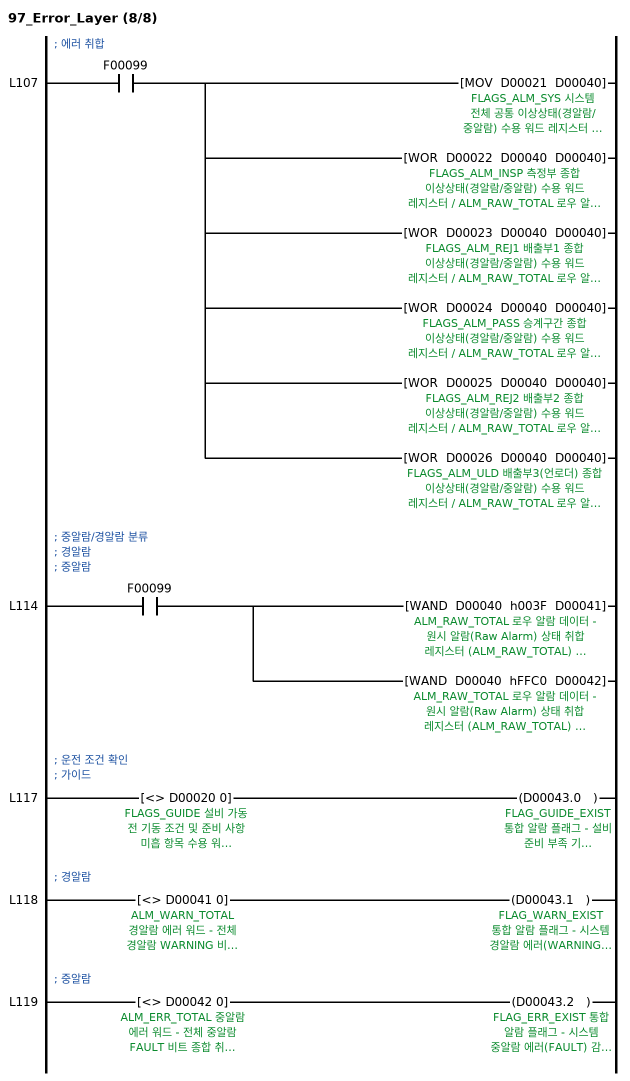
[picture p24: 97_Error_Layer rungs L107-L119]
// 에러 취합
; L107
LOAD      F00099
MOV       D00021 D00040	// FLAGS_ALM_SYS 시스템 전체 공통 이상상태(경알람/중알람) 수용 워드 레지스터 / ALM_RAW_TOTAL 로우 알람 데이터 - 원시 알람(Raw Alarm) 상태 취합 레지스터 (ALM_RAW_TOTAL)
WOR       D00022 D00040 D00040	// FLAGS_ALM_INSP 측정부 종합 이상상태(경알람/중알람) 수용 워드 레지스터 / ALM_RAW_TOTAL 로우 알람 데이터 - 원시 알람(Raw Alarm) 상태 취합 레지스터 (ALM_RAW_TOTAL) / ALM_RAW_TOTAL 로우 알람 데이터 - 원시 알람(Raw Alarm) 상태 취합 레지스터 (ALM_RAW_TOTAL)
WOR       D00023 D00040 D00040	// FLAGS_ALM_REJ1 배출부1 종합 이상상태(경알람/중알람) 수용 워드 레지스터 / ALM_RAW_TOTAL 로우 알람 데이터 - 원시 알람(Raw Alarm) 상태 취합 레지스터 (ALM_RAW_TOTAL) / ALM_RAW_TOTAL 로우 알람 데이터 - 원시 알람(Raw Alarm) 상태 취합 레지스터 (ALM_RAW_TOTAL)
WOR       D00024 D00040 D00040	// FLAGS_ALM_PASS 승계구간 종합 이상상태(경알람/중알람) 수용 워드 레지스터 / ALM_RAW_TOTAL 로우 알람 데이터 - 원시 알람(Raw Alarm) 상태 취합 레지스터 (ALM_RAW_TOTAL) / ALM_RAW_TOTAL 로우 알람 데이터 - 원시 알람(Raw Alarm) 상태 취합 레지스터 (ALM_RAW_TOTAL)
WOR       D00025 D00040 D00040	// FLAGS_ALM_REJ2 배출부2 종합 이상상태(경알람/중알람) 수용 워드 레지스터 / ALM_RAW_TOTAL 로우 알람 데이터 - 원시 알람(Raw Alarm) 상태 취합 레지스터 (ALM_RAW_TOTAL) / ALM_RAW_TOTAL 로우 알람 데이터 - 원시 알람(Raw Alarm) 상태 취합 레지스터 (ALM_RAW_TOTAL)
WOR       D00026 D00040 D00040	// FLAGS_ALM_ULD 배출부3(언로더) 종합 이상상태(경알람/중알람) 수용 워드 레지스터 / ALM_RAW_TOTAL 로우 알람 데이터 - 원시 알람(Raw Alarm) 상태 취합 레지스터 (ALM_RAW_TOTAL) / ALM_RAW_TOTAL 로우 알람 데이터 - 원시 알람(Raw Alarm) 상태 취합 레지스터 (ALM_RAW_TOTAL)
// 중알람/경알람 분류
; L114
LOAD      F00099
WAND      D00040 h003F D00041	// ALM_RAW_TOTAL 로우 알람 데이터 - 원시 알람(Raw Alarm) 상태 취합 레지스터 (ALM_RAW_TOTAL) / ALM_WARN_TOTAL 경알람 에러 워드 - 전체 경알람 WARNING 비트 종합 취합 레지스터 (ALM_WARN_TOTAL)
WAND      D00040 hFFC0 D00042	// ALM_RAW_TOTAL 로우 알람 데이터 - 원시 알람(Raw Alarm) 상태 취합 레지스터 (ALM_RAW_TOTAL) / ALM_ERR_TOTAL 중알람 에러 워드 - 전체 중알람 FAULT 비트 종합 취합 레지스터 (ALM_ERR_TOTAL)
// output comment: 경알람
// output comment: 중알람
// 운전 조건 확인
; L117
LOAD<>    D00020 0	// FLAGS_GUIDE 설비 가동 전 기동 조건 및 준비 사항 미흡 항목 수용 워드 레지스터
OUT       D00043.0	// FLAG_GUIDE_EXIST 통합 알람 플래그 - 설비 준비 부족 기동 불허(GUIDE) 활성화
// output comment: 가이드
; L118
LOAD<>    D00041 0	// ALM_WARN_TOTAL 경알람 에러 워드 - 전체 경알람 WARNING 비트 종합 취합 레지스터 (ALM_WARN_TOTAL)
OUT       D00043.1	// FLAG_WARN_EXIST 통합 알람 플래그 - 시스템 경알람 에러(WARNING) 감지 활성화
// output comment: 경알람
; L119
LOAD<>    D00042 0	// ALM_ERR_TOTAL 중알람 에러 워드 - 전체 중알람 FAULT 비트 종합 취합 레지스터 (ALM_ERR_TOTAL)
OUT       D00043.2	// FLAG_ERR_EXIST 통합 알람 플래그 - 시스템 중알람 에러(FAULT) 감지 활성화
// output comment: 중알람

PROGRAM 98_Output_Layer (task: 스캔 프로그램)

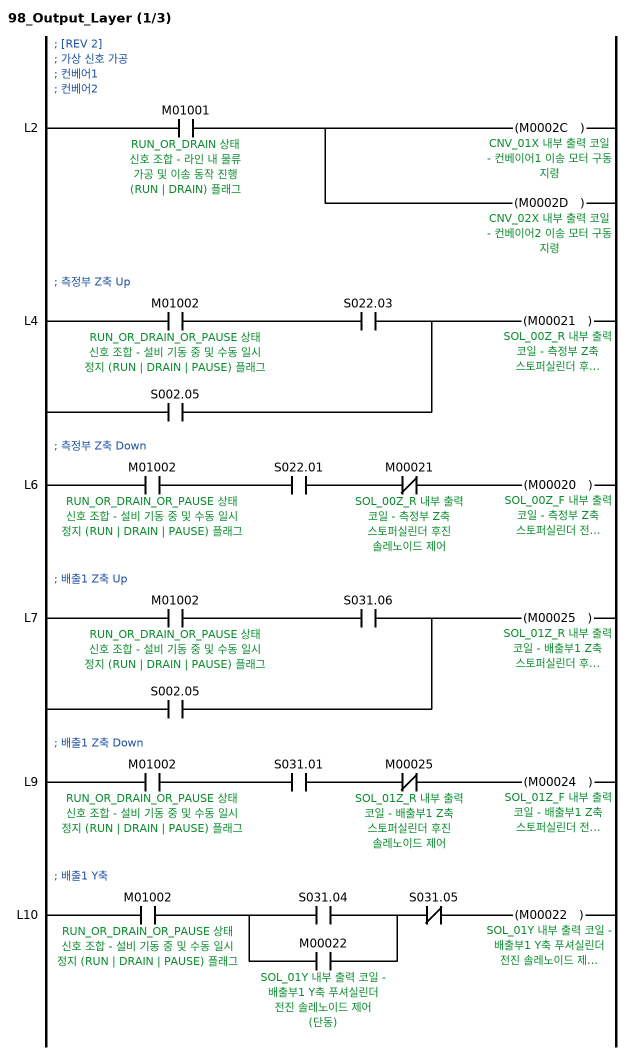
// [REV 2]
// 가상 신호 가공
; L2
LOAD      M01001	// RUN_OR_DRAIN 상태 신호 조합 - 라인 내 물류 가공 및 이송 동작 진행 (RUN | DRAIN) 플래그
OUT       M0002C	// CNV_01X 내부 출력 코일 - 컨베이어1 이송 모터 구동 지령
OUT       M0002D	// CNV_02X 내부 출력 코일 - 컨베이어2 이송 모터 구동 지령
// output comment: 컨베어1
// output comment: 컨베어2
; L4
LOAD      M01002	// RUN_OR_DRAIN_OR_PAUSE 상태 신호 조합 - 설비 기동 중 및 수동 일시 정지 (RUN | DRAIN | PAUSE) 플래그
AND       S022.03
OR        S002.05
OUT       M00021	// SOL_00Z_R 내부 출력 코일 - 측정부 Z축 스토퍼실린더 후진 솔레노이드 제어
// output comment: 측정부 Z축 Up
; L6
LOAD      M01002	// RUN_OR_DRAIN_OR_PAUSE 상태 신호 조합 - 설비 기동 중 및 수동 일시 정지 (RUN | DRAIN | PAUSE) 플래그
AND       S022.01
AND NOT   M00021	// SOL_00Z_R 내부 출력 코일 - 측정부 Z축 스토퍼실린더 후진 솔레노이드 제어
OUT       M00020	// SOL_00Z_F 내부 출력 코일 - 측정부 Z축 스토퍼실린더 전진 솔레노이드 제어
// output comment: 측정부 Z축 Down
; L7
LOAD      M01002	// RUN_OR_DRAIN_OR_PAUSE 상태 신호 조합 - 설비 기동 중 및 수동 일시 정지 (RUN | DRAIN | PAUSE) 플래그
AND       S031.06
OR        S002.05
OUT       M00025	// SOL_01Z_R 내부 출력 코일 - 배출부1 Z축 스토퍼실린더 후진 솔레노이드 제어
// output comment: 배출1 Z축 Up
; L9
LOAD      M01002	// RUN_OR_DRAIN_OR_PAUSE 상태 신호 조합 - 설비 기동 중 및 수동 일시 정지 (RUN | DRAIN | PAUSE) 플래그
AND       S031.01
AND NOT   M00025	// SOL_01Z_R 내부 출력 코일 - 배출부1 Z축 스토퍼실린더 후진 솔레노이드 제어
OUT       M00024	// SOL_01Z_F 내부 출력 코일 - 배출부1 Z축 스토퍼실린더 전진 솔레노이드 제어
// output comment: 배출1 Z축 Down
; L10
LOAD      M01002	// RUN_OR_DRAIN_OR_PAUSE 상태 신호 조합 - 설비 기동 중 및 수동 일시 정지 (RUN | DRAIN | PAUSE) 플래그
LOAD      S031.04
OR        M00022	// SOL_01Y 내부 출력 코일 - 배출부1 Y축 푸셔실린더 전진 솔레노이드 제어 (단동)
AND LOAD
AND NOT   S031.05
OUT       M00022	// SOL_01Y 내부 출력 코일 - 배출부1 Y축 푸셔실린더 전진 솔레노이드 제어 (단동)
// output comment: 배출1 Y축

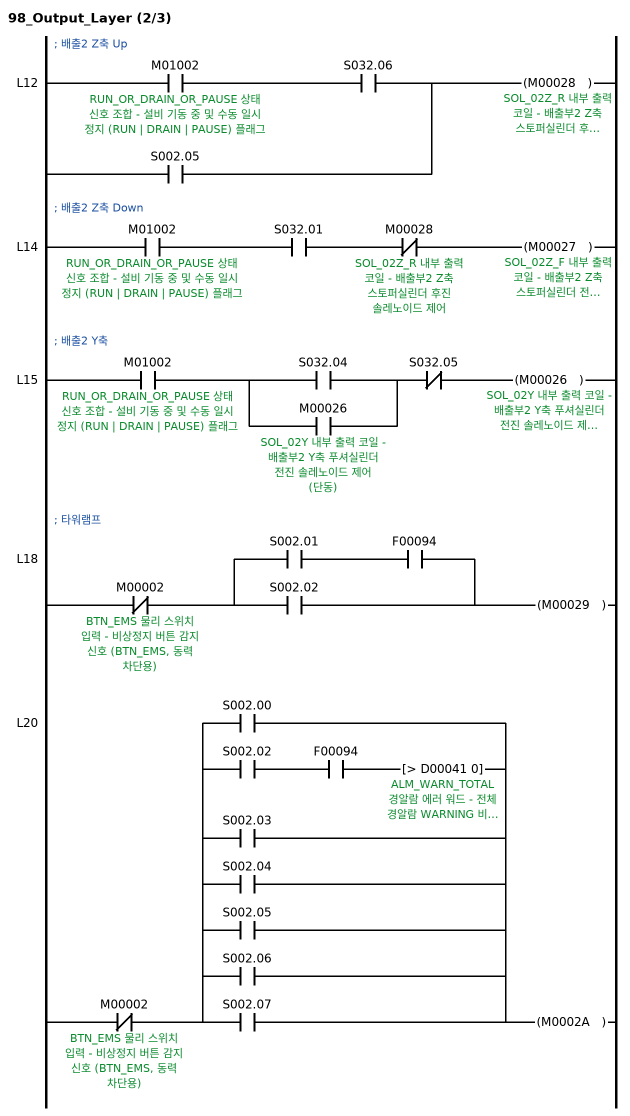
; L12
LOAD      M01002	// RUN_OR_DRAIN_OR_PAUSE 상태 신호 조합 - 설비 기동 중 및 수동 일시 정지 (RUN | DRAIN | PAUSE) 플래그
AND       S032.06
OR        S002.05
OUT       M00028	// SOL_02Z_R 내부 출력 코일 - 배출부2 Z축 스토퍼실린더 후진 솔레노이드 제어
// output comment: 배출2 Z축 Up
; L14
LOAD      M01002	// RUN_OR_DRAIN_OR_PAUSE 상태 신호 조합 - 설비 기동 중 및 수동 일시 정지 (RUN | DRAIN | PAUSE) 플래그
AND       S032.01
AND NOT   M00028	// SOL_02Z_R 내부 출력 코일 - 배출부2 Z축 스토퍼실린더 후진 솔레노이드 제어
OUT       M00027	// SOL_02Z_F 내부 출력 코일 - 배출부2 Z축 스토퍼실린더 전진 솔레노이드 제어
// output comment: 배출2 Z축 Down
; L15
LOAD      M01002	// RUN_OR_DRAIN_OR_PAUSE 상태 신호 조합 - 설비 기동 중 및 수동 일시 정지 (RUN | DRAIN | PAUSE) 플래그
LOAD      S032.04
OR        M00026	// SOL_02Y 내부 출력 코일 - 배출부2 Y축 푸셔실린더 전진 솔레노이드 제어 (단동)
AND LOAD
AND NOT   S032.05
OUT       M00026	// SOL_02Y 내부 출력 코일 - 배출부2 Y축 푸셔실린더 전진 솔레노이드 제어 (단동)
// output comment: 배출2 Y축
// 타워램프
; L18
LOAD NOT  M00002	// BTN_EMS 물리 스위치 입력 - 비상정지 버튼 감지 신호 (BTN_EMS, 동력 차단용)
LOAD      S002.01
AND       F00094
OR        S002.02
AND LOAD
OUT       M00029
; L20
LOAD NOT  M00002	// BTN_EMS 물리 스위치 입력 - 비상정지 버튼 감지 신호 (BTN_EMS, 동력 차단용)
LOAD      S002.00
LOAD      S002.02
AND       F00094
AND>      D00041 0	// ALM_WARN_TOTAL 경알람 에러 워드 - 전체 경알람 WARNING 비트 종합 취합 레지스터 (ALM_WARN_TOTAL)
OR LOAD
OR        S002.03
OR        S002.04
OR        S002.05
OR        S002.06
OR        S002.07
AND LOAD
OUT       M0002A

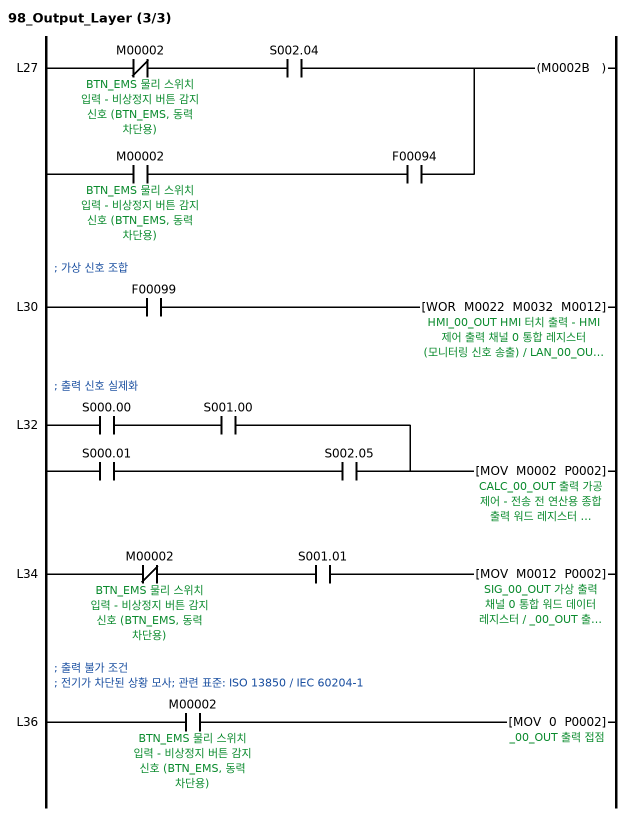
; L27
LOAD NOT  M00002	// BTN_EMS 물리 스위치 입력 - 비상정지 버튼 감지 신호 (BTN_EMS, 동력 차단용)
AND       S002.04
LOAD      M00002	// BTN_EMS 물리 스위치 입력 - 비상정지 버튼 감지 신호 (BTN_EMS, 동력 차단용)
AND       F00094
OR LOAD
OUT       M0002B
// 가상 신호 조합
; L30
LOAD      F00099
WOR       M0022 M0032 M0012	// HMI_00_OUT HMI 터치 출력 - HMI 제어 출력 채널 0 통합 레지스터 (모니터링 신호 송출) / LAN_00_OUT 통신 출력 - LAN(Modbus) 출력 채널 0 통합 레지스터 (상태 피드백 전송) / SIG_00_OUT 가상 출력 채널 0 통합 워드 데이터 레지스터
// 출력 신호 실제화
; L32
LOAD      S000.00
AND       S001.00
LOAD      S000.01
AND       S002.05
OR LOAD
MOV       M0002 P0002	// CALC_00_OUT 출력 가공 제어 - 전송 전 연산용 종합 출력 워드 레지스터 / _00_OUT 출력 접점
; L34
LOAD NOT  M00002	// BTN_EMS 물리 스위치 입력 - 비상정지 버튼 감지 신호 (BTN_EMS, 동력 차단용)
AND       S001.01
MOV       M0012 P0002	// SIG_00_OUT 가상 출력 채널 0 통합 워드 데이터 레지스터 / _00_OUT 출력 접점
// 출력 불가 조건
; L36
LOAD      M00002	// BTN_EMS 물리 스위치 입력 - 비상정지 버튼 감지 신호 (BTN_EMS, 동력 차단용)
MOV       0 P0002	// _00_OUT 출력 접점
// output comment: 전기가 차단된 상황 모사; 관련 표준: ISO 13850 / IEC 60204-1

PROGRAM 99_SubRoutine_Layer (task: 스캔 프로그램)

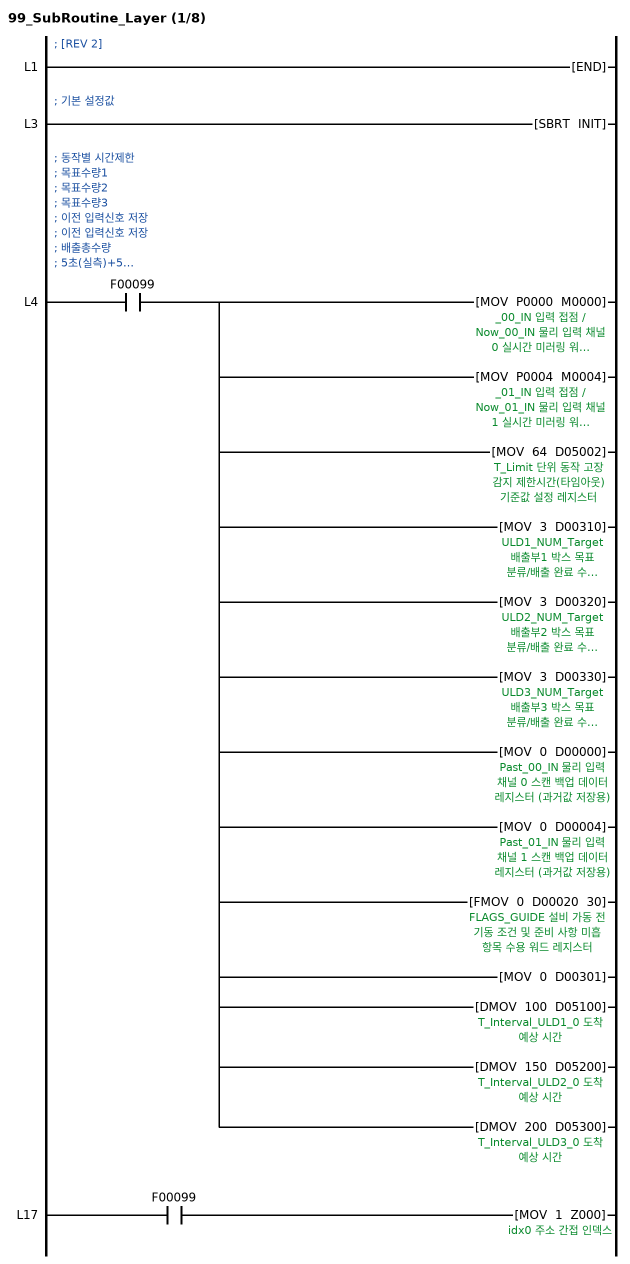
// [REV 2]
; L1
END
// 기본 설정값
; L3
SBRT      INIT
; L4
LOAD      F00099
MOV       P0000 M0000	// _00_IN 입력 접점 / Now_00_IN 물리 입력 채널 0 실시간 미러링 워드 레지스터 (Past_00_IN 비교용)
MOV       P0004 M0004	// _01_IN 입력 접점 / Now_01_IN 물리 입력 채널 1 실시간 미러링 워드 레지스터 (Past_01_IN 비교용)
MOV       64 D05002	// T_Limit 단위 동작 고장 감지 제한시간(타임아웃) 기준값 설정 레지스터
MOV       3 D00310	// ULD1_NUM_Target 배출부1 박스 목표 분류/배출 완료 수량 레지스터
MOV       3 D00320	// ULD2_NUM_Target 배출부2 박스 목표 분류/배출 완료 수량 레지스터
MOV       3 D00330	// ULD3_NUM_Target 배출부3 박스 목표 분류/배출 완료 수량 레지스터
MOV       0 D00000	// Past_00_IN 물리 입력 채널 0 스캔 백업 데이터 레지스터 (과거값 저장용)
MOV       0 D00004	// Past_01_IN 물리 입력 채널 1 스캔 백업 데이터 레지스터 (과거값 저장용)
FMOV      0 D00020 30	// FLAGS_GUIDE 설비 가동 전 기동 조건 및 준비 사항 미흡 항목 수용 워드 레지스터
MOV       0 D00301
DMOV      100 D05100	// T_Interval_ULD1_0 도착 예상 시간
DMOV      150 D05200	// T_Interval_ULD2_0 도착 예상 시간
DMOV      200 D05300	// T_Interval_ULD3_0 도착 예상 시간
// output comment: 동작별 시간제한
// output comment: 목표수량1
// output comment: 목표수량2
// output comment: 목표수량3
// output comment: 이전 입력신호 저장
// output comment: 이전 입력신호 저장
// output comment: 배출총수량
// output comment: 5초(실측)+5초
// output comment: 10초(실측)+5초
// output comment: 13초(실측)+7초
; L17
LOAD      F00099
MOV       1 Z000	// idx0 주소 간접 인덱스

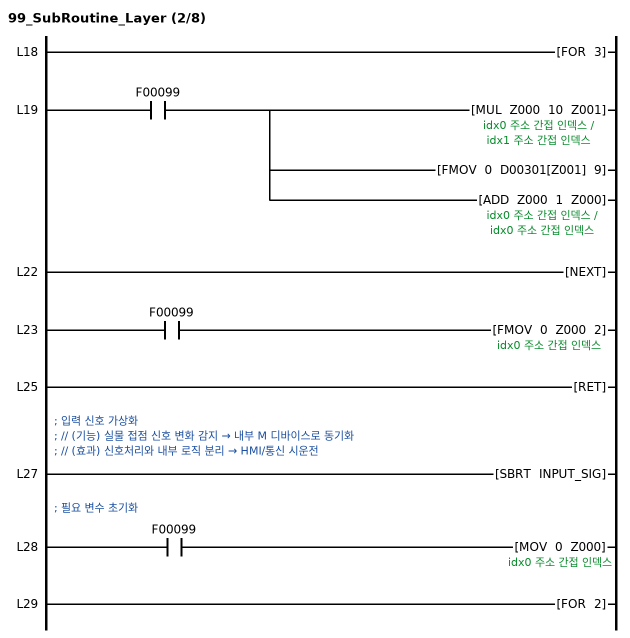
; L18
FOR       3
; L19
LOAD      F00099
MUL       Z000 10 Z001	// idx0 주소 간접 인덱스 / idx1 주소 간접 인덱스
FMOV      0 D00301[Z001] 9
ADD       Z000 1 Z000	// idx0 주소 간접 인덱스 / idx0 주소 간접 인덱스
; L22
NEXT
; L23
LOAD      F00099
FMOV      0 Z000 2	// idx0 주소 간접 인덱스
; L25
RET
// 
// 입력 신호 가상화
// // (기능) 실물 접점 신호 변화 감지 → 내부 M 디바이스로 동기화
// // (효과) 신호처리와 내부 로직 분리 → HMI/통신 시운전
; L27
SBRT      INPUT_SIG
; L28
LOAD      F00099
MOV       0 Z000	// idx0 주소 간접 인덱스
// output comment: 필요 변수 초기화
; L29
FOR       2

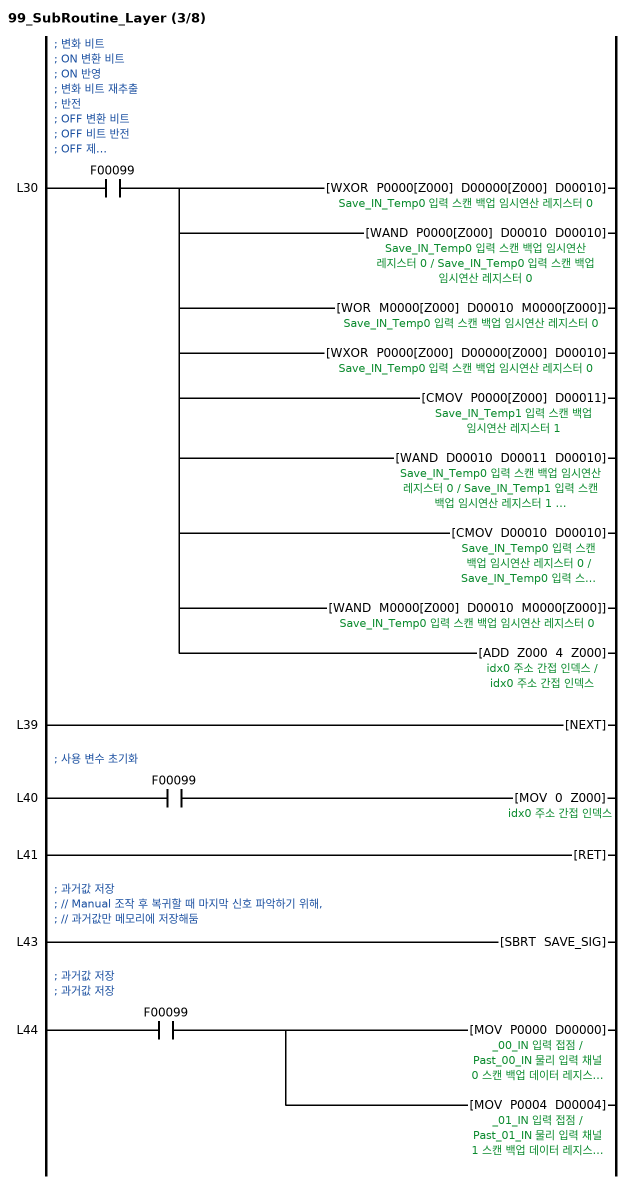
; L30
LOAD      F00099
WXOR      P0000[Z000] D00000[Z000] D00010	// Save_IN_Temp0 입력 스캔 백업 임시연산 레지스터 0
WAND      P0000[Z000] D00010 D00010	// Save_IN_Temp0 입력 스캔 백업 임시연산 레지스터 0 / Save_IN_Temp0 입력 스캔 백업 임시연산 레지스터 0
WOR       M0000[Z000] D00010 M0000[Z000]	// Save_IN_Temp0 입력 스캔 백업 임시연산 레지스터 0
WXOR      P0000[Z000] D00000[Z000] D00010	// Save_IN_Temp0 입력 스캔 백업 임시연산 레지스터 0
CMOV      P0000[Z000] D00011	// Save_IN_Temp1 입력 스캔 백업 임시연산 레지스터 1
WAND      D00010 D00011 D00010	// Save_IN_Temp0 입력 스캔 백업 임시연산 레지스터 0 / Save_IN_Temp1 입력 스캔 백업 임시연산 레지스터 1 / Save_IN_Temp0 입력 스캔 백업 임시연산 레지스터 0
CMOV      D00010 D00010	// Save_IN_Temp0 입력 스캔 백업 임시연산 레지스터 0 / Save_IN_Temp0 입력 스캔 백업 임시연산 레지스터 0
WAND      M0000[Z000] D00010 M0000[Z000]	// Save_IN_Temp0 입력 스캔 백업 임시연산 레지스터 0
ADD       Z000 4 Z000	// idx0 주소 간접 인덱스 / idx0 주소 간접 인덱스
// output comment: 변화 비트
// output comment: ON 변환 비트
// output comment: ON 반영
// output comment: 변화 비트 재추출
// output comment: 반전
// output comment: OFF 변환 비트
// output comment: OFF 비트 반전
// output comment: OFF 제거
// output comment: 40번대로 넘어감
; L39
NEXT
; L40
LOAD      F00099
MOV       0 Z000	// idx0 주소 간접 인덱스
// output comment: 사용 변수 초기화
; L41
RET
// 
// 과거값 저장
// // Manual 조작 후 복귀할 때 마지막 신호 파악하기 위해,
// // 과거값만 메모리에 저장해둠
; L43
SBRT      SAVE_SIG
; L44
LOAD      F00099
MOV       P0000 D00000	// _00_IN 입력 접점 / Past_00_IN 물리 입력 채널 0 스캔 백업 데이터 레지스터 (과거값 저장용)
MOV       P0004 D00004	// _01_IN 입력 접점 / Past_01_IN 물리 입력 채널 1 스캔 백업 데이터 레지스터 (과거값 저장용)
// output comment: 과거값 저장
// output comment: 과거값 저장

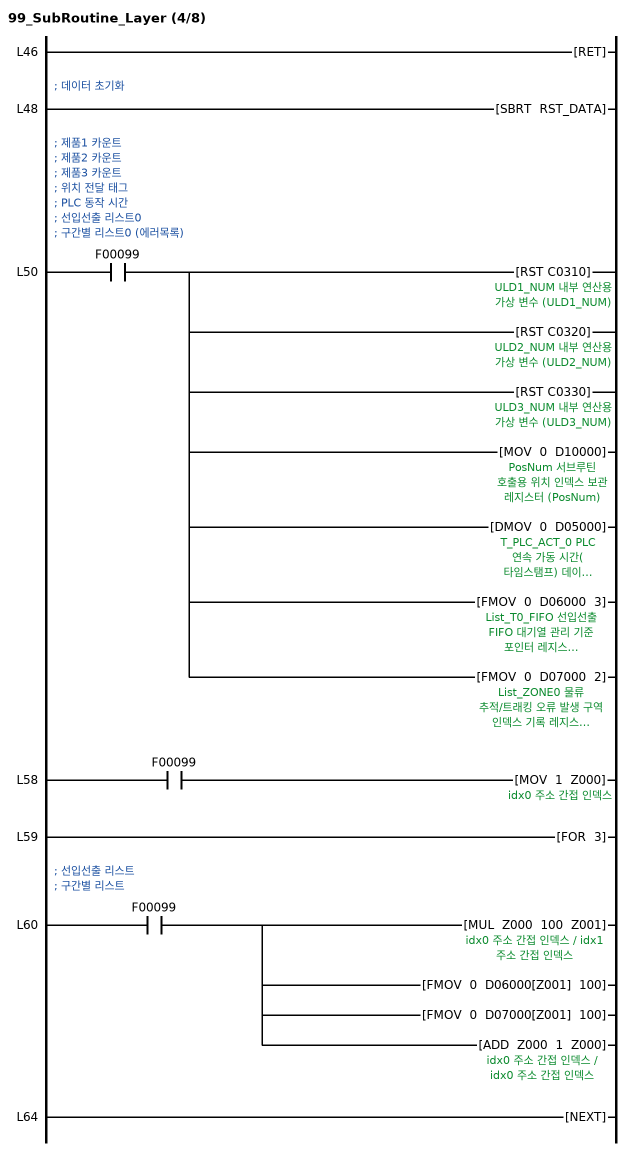
; L46
RET
// 데이터 초기화
; L48
SBRT      RST_DATA
; L50
LOAD      F00099
RST       C0310	// ULD1_NUM 내부 연산용 가상 변수 (ULD1_NUM)
RST       C0320	// ULD2_NUM 내부 연산용 가상 변수 (ULD2_NUM)
RST       C0330	// ULD3_NUM 내부 연산용 가상 변수 (ULD3_NUM)
MOV       0 D10000	// PosNum 서브루틴 호출용 위치 인덱스 보관 레지스터 (PosNum)
DMOV      0 D05000	// T_PLC_ACT_0 PLC 연속 가동 시간(타임스탬프) 데이터 레지스터 하위 16비트 (0.1초 해상도)
FMOV      0 D06000 3	// List_T0_FIFO 선입선출 FIFO 대기열 관리 기준 포인터 레지스터 (List_T0_FIFO)
FMOV      0 D07000 2	// List_ZONE0 물류 추적/트래킹 오류 발생 구역 인덱스 기록 레지스터 (List_ZONE0)
// output comment: 제품1 카운트
// output comment: 제품2 카운트
// output comment: 제품3 카운트
// output comment: 위치 전달 태그
// output comment: PLC 동작 시간
// output comment: 선입선출 리스트0
// output comment: 구간별 리스트0 (에러목록)
; L58
LOAD      F00099
MOV       1 Z000	// idx0 주소 간접 인덱스
; L59
FOR       3
; L60
LOAD      F00099
MUL       Z000 100 Z001	// idx0 주소 간접 인덱스 / idx1 주소 간접 인덱스
FMOV      0 D06000[Z001] 100
FMOV      0 D07000[Z001] 100
ADD       Z000 1 Z000	// idx0 주소 간접 인덱스 / idx0 주소 간접 인덱스
// output comment: 선입선출 리스트
// output comment: 구간별 리스트
; L64
NEXT

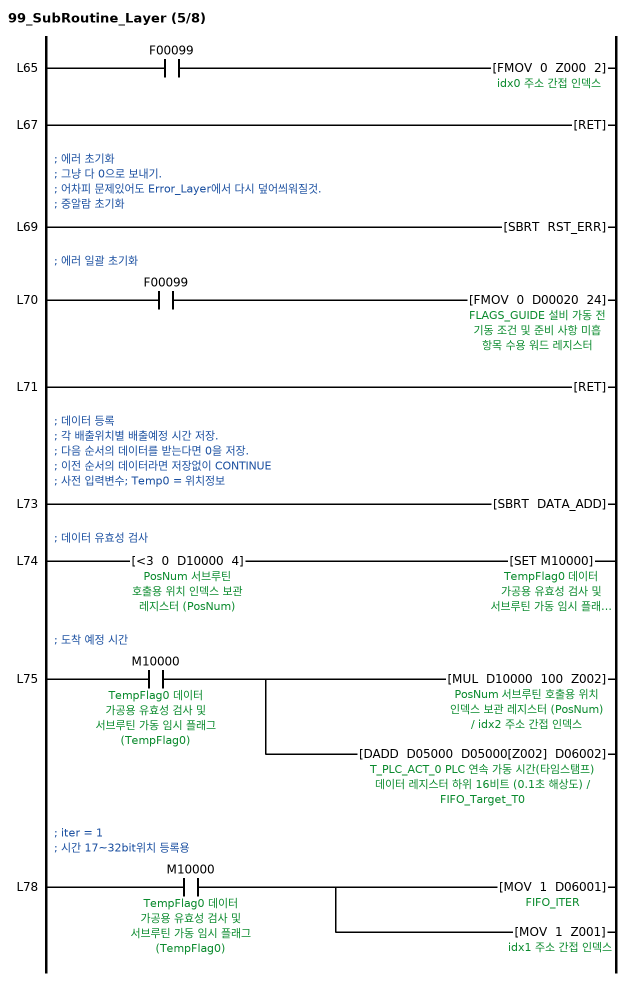
; L65
LOAD      F00099
FMOV      0 Z000 2	// idx0 주소 간접 인덱스
; L67
RET
// 
// 에러 초기화
// 
// 그냥 다 0으로 보내기.
// 어차피 문제있어도 Error_Layer에서 다시 덮어씌워질것.
; L69
SBRT      RST_ERR
// output comment: 중알람 초기화
; L70
LOAD      F00099
FMOV      0 D00020 24	// FLAGS_GUIDE 설비 가동 전 기동 조건 및 준비 사항 미흡 항목 수용 워드 레지스터
// output comment: 에러 일괄 초기화
; L71
RET
// 
// 데이터 등록
// 
// 각 배출위치별 배출예정 시간 저장.
// 다음 순서의 데이터를 받는다면 0을 저장.
// 이전 순서의 데이터라면 저장없이 CONTINUE
//  
; L73
SBRT      DATA_ADD
// output comment: 사전 입력변수; Temp0 = 위치정보
; L74
LOAD<3    0 D10000 4	// PosNum 서브루틴 호출용 위치 인덱스 보관 레지스터 (PosNum)
SET       M10000	// TempFlag0 데이터 가공용 유효성 검사 및 서브루틴 가동 임시 플래그 (TempFlag0)
// output comment: 데이터 유효성 검사
; L75
LOAD      M10000	// TempFlag0 데이터 가공용 유효성 검사 및 서브루틴 가동 임시 플래그 (TempFlag0)
MUL       D10000 100 Z002	// PosNum 서브루틴 호출용 위치 인덱스 보관 레지스터 (PosNum) / idx2 주소 간접 인덱스
DADD      D05000 D05000[Z002] D06002	// T_PLC_ACT_0 PLC 연속 가동 시간(타임스탬프) 데이터 레지스터 하위 16비트 (0.1초 해상도) / FIFO_Target_T0
// output comment: 도착 예정 시간
; L78
LOAD      M10000	// TempFlag0 데이터 가공용 유효성 검사 및 서브루틴 가동 임시 플래그 (TempFlag0)
MOV       1 D06001	// FIFO_ITER
MOV       1 Z001	// idx1 주소 간접 인덱스
// output comment: iter = 1
// output comment: 시간 17~32bit위치 등록용

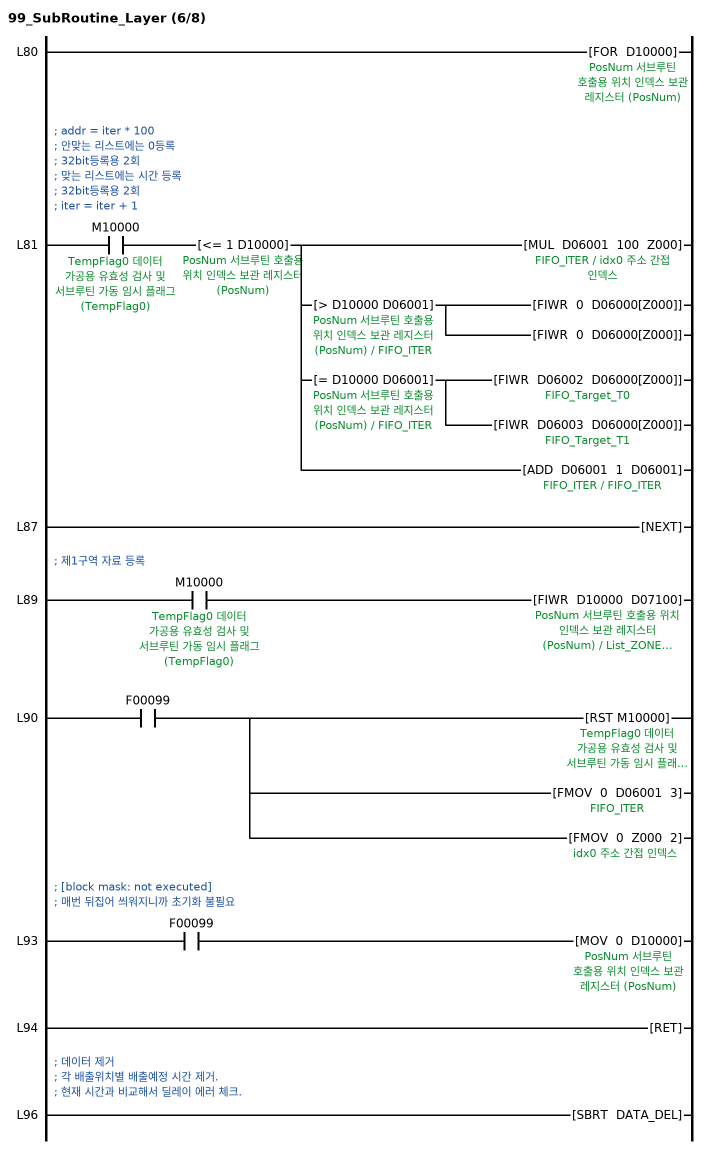
; L80
FOR       D10000	// PosNum 서브루틴 호출용 위치 인덱스 보관 레지스터 (PosNum)
; L81
LOAD      M10000	// TempFlag0 데이터 가공용 유효성 검사 및 서브루틴 가동 임시 플래그 (TempFlag0)
AND<=     1 D10000	// PosNum 서브루틴 호출용 위치 인덱스 보관 레지스터 (PosNum)
MUL       D06001 100 Z000	// FIFO_ITER / idx0 주소 간접 인덱스
MPUSH
AND>      D10000 D06001	// PosNum 서브루틴 호출용 위치 인덱스 보관 레지스터 (PosNum) / FIFO_ITER
FIWR      0 D06000[Z000]
FIWR      0 D06000[Z000]
MLOAD
AND=      D10000 D06001	// PosNum 서브루틴 호출용 위치 인덱스 보관 레지스터 (PosNum) / FIFO_ITER
FIWR      D06002 D06000[Z000]	// FIFO_Target_T0
FIWR      D06003 D06000[Z000]	// FIFO_Target_T1
MPOP
ADD       D06001 1 D06001	// FIFO_ITER / FIFO_ITER
// output comment: addr = iter * 100
// output comment: 안맞는 리스트에는 0등록
// output comment: 32bit등록용 2회
// output comment: 맞는 리스트에는 시간 등록
// output comment: 32bit등록용 2회
// output comment: iter = iter + 1
; L87
NEXT
; L89
LOAD      M10000	// TempFlag0 데이터 가공용 유효성 검사 및 서브루틴 가동 임시 플래그 (TempFlag0)
FIWR      D10000 D07100	// PosNum 서브루틴 호출용 위치 인덱스 보관 레지스터 (PosNum) / List_ZONE1 배출 영역1 물류 트래킹 데이터 적재 레지스터 (List_ZONE1)
// output comment: 제1구역 자료 등록
; L90
LOAD      F00099
RST       M10000	// TempFlag0 데이터 가공용 유효성 검사 및 서브루틴 가동 임시 플래그 (TempFlag0)
FMOV      0 D06001 3	// FIFO_ITER
FMOV      0 Z000 2	// idx0 주소 간접 인덱스
; L93 (block mask: not executed)
LOAD      F00099
MOV       0 D10000	// PosNum 서브루틴 호출용 위치 인덱스 보관 레지스터 (PosNum)
// output comment: 매번 뒤집어 씌워지니까 초기화 불필요
; L94
RET
// 
// 데이터 제거
// 
// 각 배출위치별 배출예정 시간 제거.
// 현재 시간과 비교해서 딜레이 에러 체크.
//  
; L96
SBRT      DATA_DEL

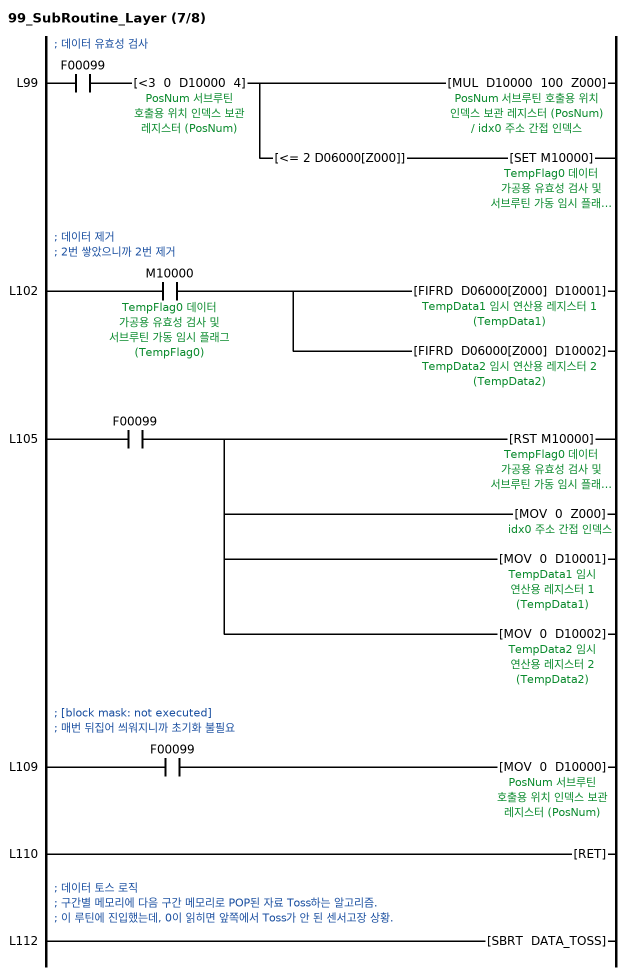
; L99
LOAD      F00099
AND<3     0 D10000 4	// PosNum 서브루틴 호출용 위치 인덱스 보관 레지스터 (PosNum)
MUL       D10000 100 Z000	// PosNum 서브루틴 호출용 위치 인덱스 보관 레지스터 (PosNum) / idx0 주소 간접 인덱스
AND<=     2 D06000[Z000]
SET       M10000	// TempFlag0 데이터 가공용 유효성 검사 및 서브루틴 가동 임시 플래그 (TempFlag0)
// output comment: 데이터 유효성 검사
; L102
LOAD      M10000	// TempFlag0 데이터 가공용 유효성 검사 및 서브루틴 가동 임시 플래그 (TempFlag0)
FIFRD     D06000[Z000] D10001	// TempData1 임시 연산용 레지스터 1 (TempData1)
FIFRD     D06000[Z000] D10002	// TempData2 임시 연산용 레지스터 2 (TempData2)
// output comment: 데이터 제거
// output comment: 2번 쌓았으니까 2번 제거
; L105
LOAD      F00099
RST       M10000	// TempFlag0 데이터 가공용 유효성 검사 및 서브루틴 가동 임시 플래그 (TempFlag0)
MOV       0 Z000	// idx0 주소 간접 인덱스
MOV       0 D10001	// TempData1 임시 연산용 레지스터 1 (TempData1)
MOV       0 D10002	// TempData2 임시 연산용 레지스터 2 (TempData2)
; L109 (block mask: not executed)
LOAD      F00099
MOV       0 D10000	// PosNum 서브루틴 호출용 위치 인덱스 보관 레지스터 (PosNum)
// output comment: 매번 뒤집어 씌워지니까 초기화 불필요
; L110
RET
// 
// 데이터 토스 로직
// 
// 구간별 메모리에 다음 구간 메모리로 POP된 자료 Toss하는 알고리즘.
// 이 루틴에 진입했는데, 0이 읽히면 앞쪽에서 Toss가 안 된 센서고장 상황.
; L112
SBRT      DATA_TOSS

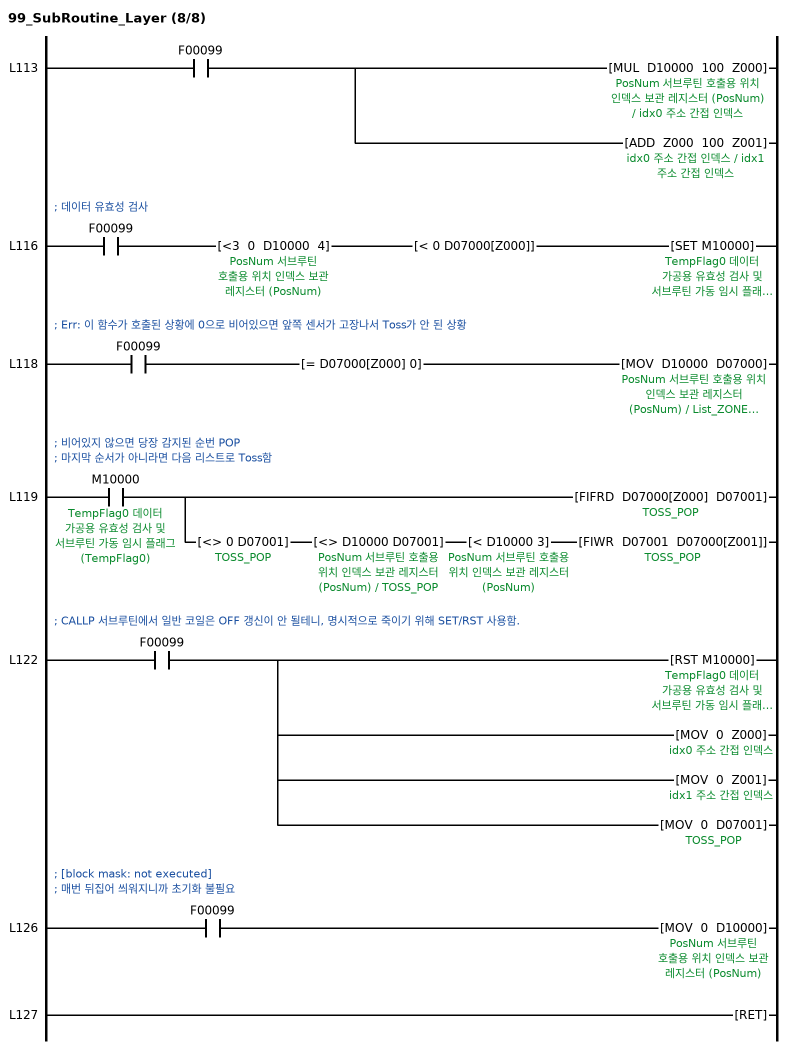
; L113
LOAD      F00099
MUL       D10000 100 Z000	// PosNum 서브루틴 호출용 위치 인덱스 보관 레지스터 (PosNum) / idx0 주소 간접 인덱스
ADD       Z000 100 Z001	// idx0 주소 간접 인덱스 / idx1 주소 간접 인덱스
; L116
LOAD      F00099
AND<3     0 D10000 4	// PosNum 서브루틴 호출용 위치 인덱스 보관 레지스터 (PosNum)
AND<      0 D07000[Z000]
SET       M10000	// TempFlag0 데이터 가공용 유효성 검사 및 서브루틴 가동 임시 플래그 (TempFlag0)
// output comment: 데이터 유효성 검사
; L118
LOAD      F00099
AND=      D07000[Z000] 0
MOV       D10000 D07000	// PosNum 서브루틴 호출용 위치 인덱스 보관 레지스터 (PosNum) / List_ZONE0 물류 추적/트래킹 오류 발생 구역 인덱스 기록 레지스터 (List_ZONE0)
// output comment: Err: 이 함수가 호출된 상황에 0으로 비어있으면 앞쪽 센서가 고장나서 Toss가 안 된 상황
; L119
LOAD      M10000	// TempFlag0 데이터 가공용 유효성 검사 및 서브루틴 가동 임시 플래그 (TempFlag0)
FIFRD     D07000[Z000] D07001	// TOSS_POP
AND<>     0 D07001	// TOSS_POP
AND<>     D10000 D07001	// PosNum 서브루틴 호출용 위치 인덱스 보관 레지스터 (PosNum) / TOSS_POP
AND<      D10000 3	// PosNum 서브루틴 호출용 위치 인덱스 보관 레지스터 (PosNum)
FIWR      D07001 D07000[Z001]	// TOSS_POP
// output comment: 비어있지 않으면 당장 감지된 순번 POP
// output comment: 마지막 순서가 아니라면 다음 리스트로 Toss함
; L122
LOAD      F00099
RST       M10000	// TempFlag0 데이터 가공용 유효성 검사 및 서브루틴 가동 임시 플래그 (TempFlag0)
MOV       0 Z000	// idx0 주소 간접 인덱스
MOV       0 Z001	// idx1 주소 간접 인덱스
MOV       0 D07001	// TOSS_POP
// output comment: CALLP 서브루틴에서 일반 코일은 OFF 갱신이 안 될테니, 명시적으로 죽이기 위해 SET/RST 사용함.
; L126 (block mask: not executed)
LOAD      F00099
MOV       0 D10000	// PosNum 서브루틴 호출용 위치 인덱스 보관 레지스터 (PosNum)
// output comment: 매번 뒤집어 씌워지니까 초기화 불필요
; L127
RET

VARIABLES AND COMMENTS (devices not used above)
D00043	WORD	ALM_SUMMARY_WORD // 통합 알람 제어 - 가이드/경알람/중알람 비트 종합 취합 레지스터 (ALM_SUMMARY_WORD)
S00100	BIT	AUTO // 전역 운전 모드 - 자동 운전 모드 (AUTO) 스텝
M00001	BIT	BTN_RUN // 물리 스위치 입력 - 자동 운전 시작 버튼 감지 신호 (BTN_RUN)
M00000	BIT	BTN_STP // 물리 스위치 입력 - 자동 운전 정지 버튼 감지 신호 (BTN_STP)
S02100	BIT	CHK_00_NA // 제품 길이 측정 완료 및 스텝 리셋 스텝
S02101	BIT	CHK_01_Length // 제품 길이 측정 시퀀스 동작 개시 및 측정 진행 스텝
S02102	BIT	CHK_02_KeepFlag // 제품 길이 측정 시퀀스 플래그값 확정
M00007	BIT	CYL_00Z_F // 물리 센서 입력 - 측정부 Z축 실린더 전진 완료 리드스위치 입력 (D-D72K)
M00008	BIT	CYL_00Z_R // 물리 센서 입력 - 측정부 Z축 실린더 후진 완료 리드스위치 입력 (D-D72K)
M00009	BIT	CYL_01Y_F // 물리 센서 입력 - 배출부1 Y축 실린더 전진 완료 리드스위치 입력 (D-D72K)
M0000A	BIT	CYL_01Y_R // 물리 센서 입력 - 배출부1 Y축 실린더 후진 완료 리드스위치 입력 (D-D72K)
M0000B	BIT	CYL_01Z_F // 물리 센서 입력 - 배출부1 Z축 실린더 전진 완료 리드스위치 입력 (D-D72K)
M0000C	BIT	CYL_01Z_R // 물리 센서 입력 - 배출부1 Z축 실린더 후진 완료 리드스위치 입력 (D-D72K)
M00040	BIT	CYL_02Y_F // 물리 센서 입력 - 배출부2 Y축 실린더 전진 완료 리드스위치 입력 (D-D72K)
M00041	BIT	CYL_02Y_R // 물리 센서 입력 - 배출부2 Y축 실린더 후진 완료 리드스위치 입력 (D-D72K)
M00042	BIT	CYL_02Z_F // 물리 센서 입력 - 배출부2 Z축 실린더 전진 완료 리드스위치 입력 (D-D72K)
M00043	BIT	CYL_02Z_R // 물리 센서 입력 - 배출부2 Z축 실린더 후진 완료 리드스위치 입력 (D-D72K)
S00001	BIT	EMERGENCY // 시스템 비상 상태 - 비상정지 스위치 활성화 (EMERGENCY) 상태 스텝
D00021.6	BIT	ERR_SYS_RESERVED_B6 // 시스템 공통 중알람 예비 비트 6
D00021.7	BIT	ERR_SYS_RESERVED_B7 // 시스템 공통 중알람 예비 비트 7
D00021.8	BIT	ERR_SYS_RESERVED_B8 // 시스템 공통 중알람 예비 비트 8
D00021.9	BIT	ERR_SYS_RESERVED_B9 // 시스템 공통 중알람 예비 비트 9
D00021.A	BIT	ERR_SYS_RESERVED_BA // 시스템 공통 중알람 예비 비트 A
D00021.B	BIT	ERR_SYS_RESERVED_BB // 시스템 공통 중알람 예비 비트 B
D00021.C	BIT	ERR_SYS_RESERVED_BC // 시스템 공통 중알람 예비 비트 C
D00021.D	BIT	ERR_SYS_RESERVED_BD // 시스템 공통 중알람 예비 비트 D
D00021.E	BIT	ERR_SYS_RESERVED_BE // 시스템 공통 중알람 예비 비트 E
D00021.F	BIT	ERR_SYS_RESERVED_BF // 시스템 공통 중알람 예비 비트 F
M00046	BIT	GET_BOX_1 // 물리 센서 입력 - 배출구1 수거박스 안착 감지 신호 (PR12-4DA 근접센서)
M00047	BIT	GET_BOX_2 // 물리 센서 입력 - 배출구2 수거박스 안착 감지 신호 (PR12-4DA 근접센서)
M00048	BIT	GET_BOX_3 // 물리 센서 입력 - 배출구3 수거박스 안착 감지 신호 (PR12-4DA 근접센서)
M00004	BIT	GET_CHK_L0 // 물리 센서 입력 - 측정부 소형 자재(길이) 감지 및 진입 판정 신호 (BYD50-DDT L0)
M00005	BIT	GET_CHK_L1 // 물리 센서 입력 - 측정부 중형 자재(길이) 감지 신호 (BYD50-DDT L1)
M00006	BIT	GET_CHK_L2 // 물리 센서 입력 - 측정부 대형 자재(길이) 감지 신호 (BYD50-DDT L2)
M0000E	BIT	GET_POS_B1 // 물리 센서 입력 - 승계구간 자재 걸림 감지 신호 (E3JK-RR12 광전센서)
M00045	BIT	GET_POS_EX // 물리 센서 입력 - 배출구3 자재 도착 감지 신호 (BY4M-PDT 광전센서)
M0000F	BIT	GET_POS_IN // 물리 센서 입력 - 측정부 자재 진입로 도착 감지 신호 (BY4M-PDT 광전센서)
M0000D	BIT	GET_POS_W1 // 물리 센서 입력 - 배출구1 자재 도착 감지 신호 (BY4M-PDT 광전센서)
M00044	BIT	GET_POS_W2 // 물리 센서 입력 - 배출구2 자재 도착 감지 신호 (BY4M-PDT 광전센서)
D00020.9	BIT	GUIDE_RESERVED_B9 // 설비 기동 가이드 예비 비트 9
D00020.A	BIT	GUIDE_RESERVED_BA // 설비 기동 가이드 예비 비트 A
D00020.B	BIT	GUIDE_RESERVED_BB // 설비 기동 가이드 예비 비트 B
D00020.C	BIT	GUIDE_RESERVED_BC // 설비 기동 가이드 예비 비트 C
D00020.D	BIT	GUIDE_RESERVED_BD // 설비 기동 가이드 예비 비트 D
D00020.E	BIT	GUIDE_RESERVED_BE // 설비 기동 가이드 예비 비트 E
D00020.F	BIT	GUIDE_RESERVED_BF // 설비 기동 가이드 예비 비트 F
S02200	BIT	LD_00_CylZDw // 측정부 배출 완료 확인 및 시퀀스 원점 복귀 종료 스텝
S02201	BIT	LD_01_GetItem // 측정부 자재 진입로 도착 감지 스텝
S02202	BIT	LD_02_CylZup // 측정부 Z축 스토퍼실린더 하강(자재 정지 및 측정 대기) 동작 스텝
S02203	BIT	LD_03_ExitItem // 측정부 제품 크기 판정 완료 및 FIFO 트래킹 데이터 등록(DATA_ADD) 스텝
S02204	BIT	LD_04_KeepUp // 측정부 Z축 스토퍼실린더 상승(자재 통과 허용) 동작 스텝
M03002	BIT	LD_QR_Err
D06102	WORD	List_T1_FIFO_1stValue_1 // 배출부1 선입선출 FIFO 도착 예정 시간 데이터 레지스터 상위 16비트 (32비트 연산)
D06202	WORD	List_T2_FIFO_1stValue_1 // 배출부2 선입선출 FIFO 도착 예정 시간 데이터 레지스터 상위 16비트 (32비트 연산)
D06302	WORD	List_T3_FIFO_1stValue_1 // 배출부3 선입선출 FIFO 도착 예정 시간 데이터 레지스터 상위 16비트 (32비트 연산)
S00101	BIT	MANUAL // 전역 운전 모드 - 수동 제어 모드 (MANUAL) 스텝
S02300	BIT	QR_00_NA
S02301	BIT	QR_01_Length
S02302	BIT	QR_02_KeepFlag
S00000	BIT	SAFE // 시스템 안전 상태 - 정상 운전 가능 (SAFE) 상태 스텝
M00102	BIT	SIG_BTN_EMS // 가상 제어 입력 - 비상정지(EMS) 활성화 통합 신호
M0012C	BIT	SIG_CNV_01X // 가상 출력 코일 - 컨베이어1 모터 기동 지령 통합 출력
M0012D	BIT	SIG_CNV_02X // 가상 출력 코일 - 컨베이어2 모터 기동 지령 통합 출력
M00120	BIT	SIG_SOL_00Z_F // 가상 출력 코일 - 측정부 Z축 스토퍼실린더 전진 솔레노이드 밸브 통합 출력
M00121	BIT	SIG_SOL_00Z_R // 가상 출력 코일 - 측정부 Z축 스토퍼실린더 후진 솔레노이드 밸브 통합 출력
M00122	BIT	SIG_SOL_01Y // 가상 출력 코일 - 배출부1 Y축 푸셔실린더 전진 솔레노이드 밸브 통합 출력 (단동)
M00124	BIT	SIG_SOL_01Z_F // 가상 출력 코일 - 배출부1 Z축 스토퍼실린더 전진 솔레노이드 밸브 통합 출력
M00125	BIT	SIG_SOL_01Z_R // 가상 출력 코일 - 배출부1 Z축 스토퍼실린더 후진 솔레노이드 밸브 통합 출력
M00126	BIT	SIG_SOL_02Y // 가상 출력 코일 - 배출부2 Y축 푸셔실린더 전진 솔레노이드 밸브 통합 출력 (단동)
M00127	BIT	SIG_SOL_02Z_F // 가상 출력 코일 - 배출부2 Z축 스토퍼실린더 전진 솔레노이드 밸브 통합 출력
M00128	BIT	SIG_SOL_02Z_R // 가상 출력 코일 - 배출부2 Z축 스토퍼실린더 후진 솔레노이드 밸브 통합 출력
S00203	BIT	STATE_DRAIN // 시스템 운전 상태 - 라인 내 잔류 물류 소진 및 정지 작업 (DRAIN) 상태 스텝
S00204	BIT	STATE_FAULT // 시스템 운전 상태 - 중알람 에러 감지 및 가동 중단 (FAULT) 상태 스텝
S00200	BIT	STATE_IDLE // 시스템 운전 상태 - 무부하 초기 대기 (IDLE) 상태 스텝
S00206	BIT	STATE_JOG // 시스템 운전 상태 - 수동 및 조그 제어 (JOG) 상태 스텝
S00207	BIT	STATE_PAUSE // 시스템 운전 상태 - 일시 정지 (PAUSE) 상태 스텝
S00201	BIT	STATE_READY // 시스템 운전 상태 - 자동 기동 조건 충족 및 대기 (READY) 상태 스텝
S00205	BIT	STATE_RESET // 시스템 운전 상태 - 원점 복귀 및 메모리 리셋 (RESET) 상태 스텝
S00202	BIT	STATE_RUN // 시스템 운전 상태 - 자동 운전 가동 (RUN) 상태 스텝
D00044	WORD	SUMMARY
D10003	WORD	TempData3 // 임시 연산용 레지스터 3 (TempData3)
D05101	WORD	T_Interval_ULD1_1 // 도착 예상 시간
D05201	WORD	T_Interval_ULD2_1 // 도착 예상 시간
D05301	WORD	T_Interval_ULD3_1 // 도착 예상 시간
D05001	WORD	T_PLC_ACT_1 // PLC 연속 가동 시간(타임스탬프) 데이터 레지스터 상위 16비트 (0.1초 해상도)
S03100	BIT	ULD1_00_CylZUp // 배출부1 Z축 스토퍼실린더 상승 완료 및 시퀀스 종료 스텝
S03101	BIT	ULD1_01_GetItem // 배출부1 도착 자재 감지 및 트래킹 데이터 판정 스텝
S03102	BIT	ULD1_02_CylZDw // 배출부1 Z축 스토퍼실린더 하강 동작 스텝
S03103	BIT	ULD1_03_KeepDw // 배출부1 Z축 스토퍼실린더 하강 및 대기 스텝
S03104	BIT	ULD1_04_SizChk // 배출부1 도착 자재 크기 재검사 및 대상 판정 스텝
S03105	BIT	ULD1_05_CylYAct // 배출부1 Y축 배출실린더 전진(제품 밀어내기 및 배출 완료 카운트) 스텝
S03106	BIT	ULD1_06_CylYBack // 배출부1 Y축 배출실린더 후진 동작 스텝
S03200	BIT	ULD2_00_CylZUp // 배출부2 Z축 스토퍼실린더 상승 완료 및 시퀀스 종료 스텝
S03201	BIT	ULD2_01_GetItem // 배출부2 도착 자재 감지 및 트래킹 데이터 판정 스텝
S03202	BIT	ULD2_02_CylZDw // 배출부2 Z축 스토퍼실린더 하강 동작 스텝
S03203	BIT	ULD2_03_KeepDw // 배출부2 Z축 스토퍼실린더 하강 및 대기 스텝
S03204	BIT	ULD2_04_SizChk // 배출부2 도착 자재 크기 재검사 및 대상 판정 스텝
S03205	BIT	ULD2_05_CylYAct // 배출부2 Y축 배출실린더 전진(제품 밀어내기 및 배출 완료 카운트) 스텝
S03206	BIT	ULD2_06_CylYBack // 배출부2 Y축 배출실린더 후진 동작 스텝
S03300	BIT	ULD3_00_NA // 배출부3 완료 및 시퀀스 종료 대기 스텝
S03301	BIT	ULD3_01_GetItem // 배출부3 자재 배출 위치 도착 감지 및 완료 대기 스텝
D00021.4	BIT	WARN_SYS_RESERVED_B4 // 시스템 공통 경알람 예비 비트 4
D00021.5	BIT	WARN_SYS_RESERVED_B5 // 시스템 공통 경알람 예비 비트 5
P00000	BIT	_00_IN00 // 입력 접점 00
P00001	BIT	_00_IN01 // 입력 접점 01
P00002	BIT	_00_IN02 // 입력 접점 02
P00003	BIT	_00_IN03 // 입력 접점 03
P00004	BIT	_00_IN04 // 입력 접점 04
P00005	BIT	_00_IN05 // 입력 접점 05
P00006	BIT	_00_IN06 // 입력 접점 06
P00007	BIT	_00_IN07 // 입력 접점 07
P00008	BIT	_00_IN08 // 입력 접점 08
P00009	BIT	_00_IN09 // 입력 접점 09
P0000A	BIT	_00_IN10 // 입력 접점 10
P0000B	BIT	_00_IN11 // 입력 접점 11
P0000C	BIT	_00_IN12 // 입력 접점 12
P0000D	BIT	_00_IN13 // 입력 접점 13
P0000E	BIT	_00_IN14 // 입력 접점 14
P0000F	BIT	_00_IN15 // 입력 접점 15
P00020	BIT	_00_OUT00 // 출력 접점 00
P00021	BIT	_00_OUT01 // 출력 접점 01
P00022	BIT	_00_OUT02 // 출력 접점 02
P00023	BIT	_00_OUT03 // 출력 접점 03
P00024	BIT	_00_OUT04 // 출력 접점 04
P00025	BIT	_00_OUT05 // 출력 접점 05
P00026	BIT	_00_OUT06 // 출력 접점 06
P00027	BIT	_00_OUT07 // 출력 접점 07
P00028	BIT	_00_OUT08 // 출력 접점 08
P00029	BIT	_00_OUT09 // 출력 접점 09
P0002A	BIT	_00_OUT10 // 출력 접점 10
P0002B	BIT	_00_OUT11 // 출력 접점 11
P0002C	BIT	_00_OUT12 // 출력 접점 12
P0002D	BIT	_00_OUT13 // 출력 접점 13
P0002E	BIT	_00_OUT14 // 출력 접점 14
P0002F	BIT	_00_OUT15 // 출력 접점 15
P00040	BIT	_01_IN00 // 입력 접점 00
P00041	BIT	_01_IN01 // 입력 접점 01
P00042	BIT	_01_IN02 // 입력 접점 02
P00043	BIT	_01_IN03 // 입력 접점 03
P00044	BIT	_01_IN04 // 입력 접점 04
P00045	BIT	_01_IN05 // 입력 접점 05
P00046	BIT	_01_IN06 // 입력 접점 06
P00047	BIT	_01_IN07 // 입력 접점 07
P00048	BIT	_01_IN08 // 입력 접점 08
P00049	BIT	_01_IN09 // 입력 접점 09
P0004A	BIT	_01_IN10 // 입력 접점 10
P0004B	BIT	_01_IN11 // 입력 접점 11
P0004C	BIT	_01_IN12 // 입력 접점 12
P0004D	BIT	_01_IN13 // 입력 접점 13
P0004E	BIT	_01_IN14 // 입력 접점 14
P0004F	BIT	_01_IN15 // 입력 접점 15